(*
SPDX-License-Identifier: MIT
License: https://opensource.org/license/mit
*)

(*!
<summary>Runs one owned multi-cycle probe for independent assertion routing.</summary>
<description>
Owns persistent root instances and fixed child storage. Use from one task without reentry.
Children borrows the same array for the instance lifetime. Root parents remain zero.
</description>
*)

{attribute 'no_assign'}
{attribute 'no_explicit_call' := 'do not call this function block directly'}
FUNCTION_BLOCK IsolationTestRunner EXTENDS TOF_Testing.TestRunner<1>
VAR_STAT
	//! <summary>Class name shared by instances of this concrete runner.</summary>
	{attribute 'hide'}
	_ClassName : STRING := __POUNAME();
END_VAR
VAR
	{attribute 'hide'}
	{attribute 'init_namespace'}
	_NamespaceName : STRING;
END_VAR
VAR_OUTPUT
	//! <summary>Owned root element used by this runner.</summary>
	Child : AssertionIsolationProbe(name := "Receiver", parent := 0);
END_VAR
VAR
	_Children : ARRAY [0.._ChildCount - 1] OF TOF_Testing.ITestElement :=
	[
		Child
	];
END_VAR

(*!
<summary>Borrows the concrete class name; callers must not modify the returned storage.</summary>
*)
{attribute 'monitoring' := 'call'}
PROPERTY ClassName : REFERENCE TO STRING
GET
ClassName REF= _ClassName;
END_GET
END_PROPERTY

(*!
<summary>Borrows the concrete namespace name for the instance lifetime; callers must not modify it.</summary>
*)
{attribute 'monitoring' := 'call'}
PROPERTY NamespaceName : REFERENCE TO STRING
GET
NamespaceName REF= _NamespaceName;
END_GET
END_PROPERTY

(*!
<summary>Reports the complete concrete instance size.</summary>
*)
{attribute 'monitoring' := 'call'}
PROPERTY SelfSize : ULINT
GET
SelfSize := XSIZEOF(THIS^);
END_GET
END_PROPERTY

(*!
<summary>Borrows the unchanged persistent root array; application code must not modify it.</summary>
*)
{attribute 'monitoring' := 'call'}
PROPERTY Children : REFERENCE TO ARRAY [0.._ChildCount - 1] OF TOF_Testing.ITestElement
GET
Children REF= _Children;
END_GET
END_PROPERTY

END_FUNCTION_BLOCK

(* stored: Version 1.1.0.1
   POU IsolationTestRunner: Id {d4040b91-f1f9-47ab-b7f5-287b0dff494a}, SpecialFunc None
   Property ClassName: Id {ffa86613-c8e3-4f6b-9dd8-097dd7819ae5}
   Get Get: Id {917aae50-ae2b-4fec-be69-d7d8b1435742}
   Property NamespaceName: Id {202be9a7-1a0e-4229-998b-7f7eed760840}
   Get Get: Id {ae483395-77ae-43ff-86b8-90f0a99011cc}
   Property SelfSize: Id {67a24499-1ec0-4e37-9d8a-4a05bdb88f5f}
   Get Get: Id {87e88cac-461c-4083-adba-ad1425ab64a6}
   Property Children: Id {70beb902-27d3-49d4-be48-461afd156f65}
   Get Get: Id {f0f48fcc-44fe-40aa-a225-6afaf668a604} *)
